ABB RAPID module: ExpProg2.mod

%%%
  VERSION:1
  LANGUAGE:ENGLISH
%%%
MODULE MOD_ExpProg2

    ! -------------------------------
    ! Define customized variables here
    ! ...

	! Tool variables:

	! Reference variables:
	PERS wobjdata F1 := [FALSE, TRUE, "", [[0,0,0],[1,0,0,0]],[[0.000,1000.000,0.000],[1.00000000,0.00000000,0.00000000,0.00000000]]];

	PROC Main()
		ConfJ \On;
		ConfL \Off;
		! Program generated by RoboDK v6.0.7 for ABB IRB 120-3/0.6 on XX/XX/XXXX 12:34:41
		! Using nominal kinematics.
		MoveAbsJ [[0.000000,-10.000000,20.000000,0.000000,30.000000,-0.000000],[9E+09,9E+09,9E+09,9E+09,9E+09,9E+09]],v500,z1,tool0 \WObj:=F1;
	ENDPROC

ENDMODULE
